{attribute 'qualified_only'}
{attribute 'strict'}
{attribute 'to_string'}
TYPE eShutterStateType :
(
    IDLE,            // Not moving
    OPENING,       // Moving upward (opening)
    CLOSING      // Moving downward (closing)
);
END_TYPE

(* stored: Version 1.1.0.1
   DUT eShutterStateType: Id {739f3d94-17ed-4c90-bd16-9c7cc9683f6f} *)
